Staubli VAL3: MatrixLib.pjx

--- MatrixLib.pjx ---
Parameters version=s8.8.3Cs9_BS1660 stackSize=5000 millimeterUnit=true
Program file=Atan2.pgx
Program file=InverseMatrix.pgx
Program file=Matrix2Trsf.pgx
Program file=MutliMatrix.pgx
Program file=Point2Trsf.pgx
Program file=Trsf2Matrix.pgx
Data file=MatrixLib.dtx

--- MatrixLib.dtx ---


--- Atan2.pgx ---
public program Atan2(num y, num x, num& angle)
begin
  //双变量反正切函数atan2(x,y)
  if x>0
    angle=atan(y/x)
  elseIf y>=0 and x<0
    angle=atan(y/x)+180
  elseIf y<0 and x<0
    angle=atan(y/x)-180
  elseIf y>0 and x==0
    angle=90
  elseIf y<0 and x==0
    angle=-90
  elseIf y==0 and x==0
    //Undefined
  endIf
end

--- InverseMatrix.pgx ---
public program InverseMatrix(num& x_nMatrixOrigin[] (dimensions=2), num& x_nMatrixNew[] (dimensions=2), bool& x_bStatus)
  local num A11
  local num A12
  local num A13
  local num A14
  local num A21
  local num A22
  local num A23
  local num A24
  local num A31
  local num A32
  local num A33
  local num A34
  local num A41
  local num A42
  local num A43
  local num A44
  local num a11
  local num a12
  local num a13
  local num a14
  local num a21
  local num a22
  local num a23
  local num a24
  local num a31
  local num a32
  local num a33
  local num a34
  local num a41
  local num a42
  local num a43
  local num a44
  local num i
  local num j
  local num A
begin
  //初始化变量
  a11=x_nMatrixOrigin[0,0]
  a21=x_nMatrixOrigin[0,1]
  a31=x_nMatrixOrigin[0,2]
  a41=x_nMatrixOrigin[0,3]
  a12=x_nMatrixOrigin[1,0]
  a22=x_nMatrixOrigin[1,1]
  a32=x_nMatrixOrigin[1,2]
  a42=x_nMatrixOrigin[1,3]
  a13=x_nMatrixOrigin[2,0]
  a23=x_nMatrixOrigin[2,1]
  a33=x_nMatrixOrigin[2,2]
  a43=x_nMatrixOrigin[2,3]
  a14=x_nMatrixOrigin[3,0]
  a24=x_nMatrixOrigin[3,1]
  a34=x_nMatrixOrigin[3,2]
  a44=x_nMatrixOrigin[3,3]

  //求代数余子式
  A11=power(-1,1+1)*(a22*a33*a44+a23*a34*a42+a24*a32*a43-a22*a34*a43-a23*a32*a44-a24*a33*a42)
  A12=power(-1,1+2)*(a21*a33*a44+a23*a34*a41+a24*a31*a43-a21*a34*a43-a23*a31*a44-a24*a33*a41)
  A13=power(-1,1+3)*(a21*a32*a44+a22*a34*a41+a24*a31*a42-a21*a34*a42-a22*a31*a44-a24*a32*a41)
  A14=power(-1,1+4)*(a21*a32*a43+a22*a33*a41+a23*a31*a42-a21*a33*a42-a22*a31*a43-a23*a32*a41)
  //
  A21=power(-1,2+1)*(a12*a33*a44+a13*a34*a42+a14*a32*a43-a12*a34*a43-a13*a32*a44-a14*a33*a42)
  A22=power(-1,2+2)*(a11*a33*a44+a13*a34*a41+a14*a31*a43-a11*a34*a43-a13*a31*a44-a14*a33*a41)
  A23=power(-1,2+3)*(a11*a32*a44+a12*a34*a41+a14*a31*a42-a11*a34*a42-a12*a31*a44-a14*a32*a41)
  A24=power(-1,2+4)*(a11*a32*a43+a12*a33*a41+a13*a31*a42-a11*a33*a42-a12*a31*a43-a13*a32*a41)
  //
  A31=power(-1,3+1)*(a12*a23*a44+a13*a24*a42+a14*a22*a43-a12*a24*a43-a13*a22*a44-a14*a23*a42)
  A32=power(-1,3+2)*(a11*a23*a44+a13*a24*a41+a14*a21*a43-a11*a24*a43-a13*a21*a44-a14*a23*a41)
  A33=power(-1,3+3)*(a11*a22*a44+a12*a24*a41+a14*a21*a42-a11*a24*a42-a12*a21*a44-a14*a22*a41)
  A34=power(-1,3+4)*(a11*a22*a43+a12*a23*a41+a13*a21*a42-a11*a23*a42-a12*a21*a43-a13*a22*a41)
  //
  A41=power(-1,4+1)*(a12*a23*a34+a13*a24*a32+a14*a22*a33-a12*a24*a33-a13*a22*a34-a14*a23*a32)
  A42=power(-1,4+2)*(a11*a23*a34+a13*a24*a31+a14*a21*a33-a11*a24*a33-a13*a21*a34-a14*a23*a31)
  A43=power(-1,4+3)*(a11*a22*a34+a12*a24*a31+a14*a21*a32-a11*a24*a32-a12*a21*a34-a14*a22*a31)
  A44=power(-1,4+4)*(a11*a22*a33+a12*a23*a31+a13*a21*a32-a11*a23*a32-a12*a21*a33-a13*a22*a31)

  //求行列式的值
  A=a11*A11+a12*A12+a13*A13+a14*A14


  if abs(A)<0.001
    //逆矩阵不存在
    x_bStatus=false
    for i=0 to 3
      for j=0 to 3
        x_nMatrixNew[i,j]=0
      endFor
    endFor
  else
    //逆矩阵存在
    x_bStatus=true
    x_nMatrixNew[0,0]=A11/A
    x_nMatrixNew[0,1]=A12/A
    x_nMatrixNew[0,2]=A13/A
    x_nMatrixNew[0,3]=A14/A
    x_nMatrixNew[1,0]=A21/A
    x_nMatrixNew[1,1]=A22/A
    x_nMatrixNew[1,2]=A23/A
    x_nMatrixNew[1,3]=A24/A
    x_nMatrixNew[2,0]=A31/A
    x_nMatrixNew[2,1]=A32/A
    x_nMatrixNew[2,2]=A33/A
    x_nMatrixNew[2,3]=A34/A
    x_nMatrixNew[3,0]=A41/A
    x_nMatrixNew[3,1]=A42/A
    x_nMatrixNew[3,2]=A43/A
    x_nMatrixNew[3,3]=A44/A
  endIf
end

--- Matrix2Trsf.pgx ---
public program Matrix2Trsf(num& x_nMatrix[] (dimensions=2), trsf& x_trTrsf)
  local num ax
  local num ay
  local num az
  local num nx
  local num ny
  local num nz
  local num ox
  local num oy
  local num oz
  local num px
  local num py
  local num pz
  local num rx1
  local num rx2
  local num ry1
  local num ry2
  local num rz1
  local num rz2
  local num x
  local num y
  local num z
begin
  //Matrik转换成Trsf
  nx=x_nMatrix[0,0]
  ny=x_nMatrix[0,1]
  nz=x_nMatrix[0,2]
  ox=x_nMatrix[1,0]
  oy=x_nMatrix[1,1]
  oz=x_nMatrix[1,2]
  ax=x_nMatrix[2,0]
  ay=x_nMatrix[2,1]
  az=x_nMatrix[2,2]
  px=x_nMatrix[3,0]
  py=x_nMatrix[3,1]
  pz=x_nMatrix[3,2]
  //求解Rx、Ry、Rz
  x_trTrsf.x=px
  x_trTrsf.y=py
  x_trTrsf.z=pz
  //求解Rx、Ry、Rz
  call Atan2(ax,sqrt(power(nx,2)+power(ox,2)),ry1)
  if ry1==90
    rx1=0
    call Atan2(ny,-nz,rz1)
  elseIf ry1==-90
    rx1=0
    call Atan2(ny,nz,rz1)
  else
    call Atan2(-ay/cos(ry1),az/cos(ry1),rx1)
    call Atan2(-ox/cos(ry1),nx/cos(ry1),rz1)
  endIf

  call Atan2(ax,sqrt(power(nx,2)+power(ox,2)),ry2)
  if ry2==90
    rx2=0
    call Atan2(ny,-nz,rz2)
  elseIf ry2==-90
    rx2=0
    call Atan2(ny,nz,rz2)
  else
    call Atan2(-ay/cos(ry2),az/cos(ry2),rx2)
    call Atan2(-ox/cos(ry2),nx/cos(ry2),rz2)
  endIf

  if abs(rx1)+abs(ry1)+abs(rz1)<=abs(rx2)+abs(ry2)+abs(rz2)
    x_trTrsf.rx=rx1
    x_trTrsf.ry=ry1
    x_trTrsf.rz=rz1
  else
    x_trTrsf.rx=rx2
    x_trTrsf.ry=ry2
    x_trTrsf.rz=rz2
  endIf
end

--- MutliMatrix.pgx ---
public program MutliMatrix(num& x_nMatrix1[] (dimensions=2), num& x_nMatrix2[] (dimensions=2), num& x_nMatrix3[] (dimensions=2))
  local num a11
  local num a12
  local num a13
  local num a14
  local num a21
  local num a22
  local num a23
  local num a24
  local num a31
  local num a32
  local num a33
  local num a34
  local num a41
  local num a42
  local num a43
  local num a44
  local num b11
  local num b12
  local num b13
  local num b14
  local num b21
  local num b22
  local num b23
  local num b24
  local num b31
  local num b32
  local num b33
  local num b34
  local num b41
  local num b42
  local num b43
  local num b44
begin
  //初始化变量
  a11=x_nMatrix1[0,0]
  a21=x_nMatrix1[0,1]
  a31=x_nMatrix1[0,2]
  a41=x_nMatrix1[0,3]
  a12=x_nMatrix1[1,0]
  a22=x_nMatrix1[1,1]
  a32=x_nMatrix1[1,2]
  a42=x_nMatrix1[1,3]
  a13=x_nMatrix1[2,0]
  a23=x_nMatrix1[2,1]
  a33=x_nMatrix1[2,2]
  a43=x_nMatrix1[2,3]
  a14=x_nMatrix1[3,0]
  a24=x_nMatrix1[3,1]
  a34=x_nMatrix1[3,2]
  a44=x_nMatrix1[3,3]

  b11=x_nMatrix2[0,0]
  b21=x_nMatrix2[0,1]
  b31=x_nMatrix2[0,2]
  b41=x_nMatrix2[0,3]
  b12=x_nMatrix2[1,0]
  b22=x_nMatrix2[1,1]
  b32=x_nMatrix2[1,2]
  b42=x_nMatrix2[1,3]
  b13=x_nMatrix2[2,0]
  b23=x_nMatrix2[2,1]
  b33=x_nMatrix2[2,2]
  b43=x_nMatrix2[2,3]
  b14=x_nMatrix2[3,0]
  b24=x_nMatrix2[3,1]
  b34=x_nMatrix2[3,2]
  b44=x_nMatrix2[3,3]

  //矩阵相乘

  x_nMatrix3[0,0]=a11*b11+a12*b21+a13*b31+a14*b41
  x_nMatrix3[0,1]=a21*b11+a22*b21+a23*b31+a24*b41
  x_nMatrix3[0,2]=a31*b11+a32*b21+a33*b31+a34*b41
  x_nMatrix3[0,3]=a41*b11+a42*b21+a43*b31+a44*b41

  x_nMatrix3[1,0]=a11*b12+a12*b22+a13*b32+a14*b42
  x_nMatrix3[1,1]=a21*b12+a22*b22+a23*b32+a24*b42
  x_nMatrix3[1,2]=a31*b12+a32*b22+a33*b32+a34*b42
  x_nMatrix3[1,3]=a41*b12+a42*b22+a43*b32+a44*b42

  x_nMatrix3[2,0]=a11*b13+a12*b23+a13*b33+a14*b43
  x_nMatrix3[2,1]=a21*b13+a22*b23+a23*b33+a24*b43
  x_nMatrix3[2,2]=a31*b13+a32*b23+a33*b33+a34*b43
  x_nMatrix3[2,3]=a41*b13+a42*b23+a43*b33+a44*b43

  x_nMatrix3[3,0]=a11*b14+a12*b24+a13*b34+a14*b44
  x_nMatrix3[3,1]=a21*b14+a22*b24+a23*b34+a24*b44
  x_nMatrix3[3,2]=a31*b14+a32*b24+a33*b34+a34*b44
  x_nMatrix3[3,3]=a41*b14+a42*b24+a43*b34+a44*b44
end

--- Point2Trsf.pgx ---
public program Point2Trsf(point x_pPoint, trsf& x_trTrsf)
begin
  x_trTrsf.x=x_pPoint.trsf.x
  x_trTrsf.y=x_pPoint.trsf.y
  x_trTrsf.z=x_pPoint.trsf.z
  x_trTrsf.rx=x_pPoint.trsf.rx
  x_trTrsf.ry=x_pPoint.trsf.ry
  x_trTrsf.rz=x_pPoint.trsf.rz
end

--- Trsf2Matrix.pgx ---
public program Trsf2Matrix(trsf x_trTrsf, num& x_nMatrix[] (dimensions=2))
  local num ax
  local num ay
  local num az
  local num nx
  local num ny
  local num nz
  local num ox
  local num oy
  local num oz
  local num px
  local num py
  local num pz
  local num rx
  local num ry
  local num rz
  local num x
  local num y
  local num z
begin
  //Trsf转换成Matrik
  x=x_trTrsf.x
  y=x_trTrsf.y
  z=x_trTrsf.z
  rx=x_trTrsf.rx
  ry=x_trTrsf.ry
  rz=x_trTrsf.rz
  //
  nx=cos(ry)*cos(rz)
  ny=sin(rx)*sin(ry)*cos(rz)+cos(rx)*sin(rz)
  nz=-cos(rx)*sin(ry)*cos(rz)+sin(rx)*sin(rz)
  ox=-cos(ry)*sin(rz)
  oy=-sin(rx)*sin(ry)*sin(rz)+cos(rx)*cos(rz)
  oz=cos(rx)*sin(ry)*sin(rz)+sin(rx)*cos(rz)
  ax=sin(ry)
  ay=-sin(rx)*cos(ry)
  az=cos(rx)*cos(ry)
  px=x
  py=y
  pz=z
  //
  x_nMatrix[0,0]=nx
  x_nMatrix[0,1]=ny
  x_nMatrix[0,2]=nz
  x_nMatrix[0,3]=0
  x_nMatrix[1,0]=ox
  x_nMatrix[1,1]=oy
  x_nMatrix[1,2]=oz
  x_nMatrix[1,3]=0
  x_nMatrix[2,0]=ax
  x_nMatrix[2,1]=ay
  x_nMatrix[2,2]=az
  x_nMatrix[2,3]=0
  x_nMatrix[3,0]=px
  x_nMatrix[3,1]=py
  x_nMatrix[3,2]=pz
  x_nMatrix[3,3]=1
end
